(* IEC 61131-3 sources: plc-iiot-stack/src/POUs/Iiot/F_IiotAlarmPriorityText, 2 files *)

(* ---- F_IiotAlarmPriorityText.decl.st ---- *)
// Назначение: имя приоритета тревоги для поля priority (None — пусто: тревога не
//             публикуется).
// Автор:      kr0nsch
// Версия:     0.1.0
// Документ:   docs/plc_mqtt.md, раздел «Тревоги»
FUNCTION F_IiotAlarmPriorityText : STRING(GVL_Const.IIOT_TEXT_LEN)
VAR_INPUT
    ePriority : E_IiotAlarmPriority;
END_VAR

(* ---- F_IiotAlarmPriorityText.impl.st ---- *)
CASE ePriority OF
    E_IiotAlarmPriority.Low:
        F_IiotAlarmPriorityText := 'Low';
    E_IiotAlarmPriority.Medium:
        F_IiotAlarmPriorityText := 'Medium';
    E_IiotAlarmPriority.High:
        F_IiotAlarmPriorityText := 'High';
    E_IiotAlarmPriority.Critical:
        F_IiotAlarmPriorityText := 'Critical';
ELSE
    F_IiotAlarmPriorityText := '';
END_CASE
